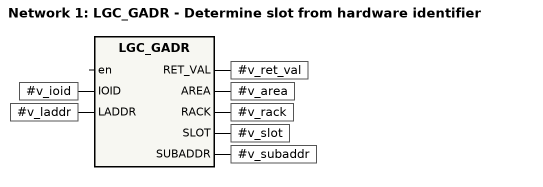
   #v_ret_val := LGC_GADR(IOID := #v_ioid,
                          LADDR := #v_laddr,
                          AREA => #v_area,
                          RACK => #v_rack,
                          SLOT => #v_slot,
                          SUBADDR => #v_subaddr);
END_REGION
END_FUNCTION_BLOCK

FUNCTION_BLOCK "FB_Fbd_ou001"   // FB169, FBD
{ S7_Optimized_Access := 'TRUE' }
   VAR_INPUT
      v_req : Bool;
      v_cont : Bool;
      v_len : UInt;
   END_VAR
   VAR_OUTPUT
      v_done : Bool;
      v_busy : Bool;
      v_error : Bool;
      v_status : Word;
   END_VAR
   VAR_IN_OUT
      v_connect : TCON_Param;
      v_data : Array[0..99] of Byte;
      v_com_rst : Bool;
      v_addr : Variant;
   END_VAR
   VAR
      inst : TSEND_C;
   END_VAR
BEGIN

REGION Network 1: TSEND_C - Send data via Ethernet
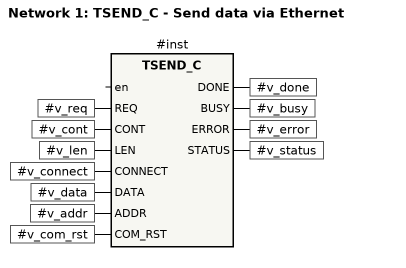
   #inst(REQ := #v_req,   // TSEND_C
         CONT := #v_cont,
         LEN := #v_len,
         CONNECT := #v_connect,
         DATA := #v_data,
         ADDR := #v_addr,
         COM_RST := #v_com_rst,
         DONE => #v_done,
         BUSY => #v_busy,
         ERROR => #v_error,
         STATUS => #v_status);
END_REGION
END_FUNCTION_BLOCK

FUNCTION_BLOCK "FB_Fbd_ou002"   // FB170, FBD
{ S7_Optimized_Access := 'TRUE' }
   VAR_INPUT
      v_req : Bool;
      v_cont : Bool;
      v_len : UDInt;
   END_VAR
   VAR_OUTPUT
      v_done : Bool;
      v_busy : Bool;
      v_error : Bool;
      v_status : Word;
   END_VAR
   VAR_IN_OUT
      v_connect : Array[0..99] of Byte;
      v_data : Array[0..99] of Byte;
      v_addr : Array[0..99] of Byte;
      v_com_rst : Bool;
   END_VAR
   VAR
      inst : TSEND_C;
   END_VAR
BEGIN

REGION Network 1: TSEND_C - Establishing a connection and sending data
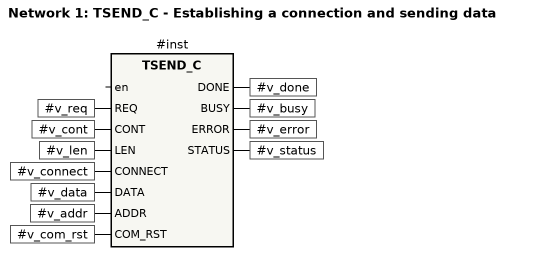
   #inst(REQ := #v_req,   // TSEND_C
         CONT := #v_cont,
         LEN := #v_len,
         CONNECT := #v_connect,
         DATA := #v_data,
         ADDR := #v_addr,
         COM_RST := #v_com_rst,
         DONE => #v_done,
         BUSY => #v_busy,
         ERROR => #v_error,
         STATUS => #v_status);
END_REGION
END_FUNCTION_BLOCK

FUNCTION_BLOCK "FB_Fbd_ou004"   // FB171, FBD
{ S7_Optimized_Access := 'TRUE' }
   VAR_INPUT
      v_en_r : Bool;
      v_cont : Bool;
      v_len : UDInt;
      v_adhoc : Bool;
   END_VAR
   VAR_OUTPUT
      v_done : Bool;
      v_busy : Bool;
      v_error : Bool;
      v_status : Word;
      v_rcvd_len : UDInt;
   END_VAR
   VAR_IN_OUT
      v_connect : Array[0..99] of Byte;
      v_data : Array[0..99] of Byte;
      v_addr : Array[0..99] of Byte;
      v_com_rst : Bool;
   END_VAR
   VAR
      inst : TRCV_C;
   END_VAR
BEGIN

REGION Network 1: TRCV_C - Establishing a connection and receiving data
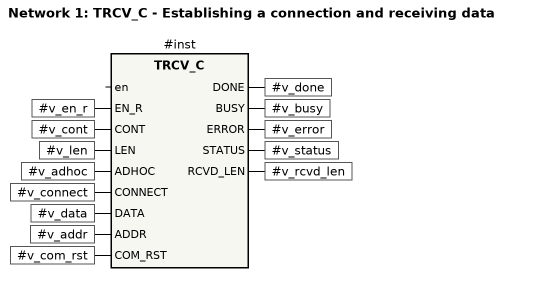
   #inst(EN_R := #v_en_r,   // TRCV_C
         CONT := #v_cont,
         LEN := #v_len,
         ADHOC := #v_adhoc,
         CONNECT := #v_connect,
         DATA := #v_data,
         ADDR := #v_addr,
         COM_RST := #v_com_rst,
         DONE => #v_done,
         BUSY => #v_busy,
         ERROR => #v_error,
         STATUS => #v_status,
         RCVD_LEN => #v_rcvd_len);
END_REGION
END_FUNCTION_BLOCK

FUNCTION_BLOCK "FB_Fbd_ou010"   // FB172, FBD
{ S7_Optimized_Access := 'TRUE' }
   VAR_INPUT
      v_req : Bool;
      v_id : Conn_Ouc;
   END_VAR
   VAR_OUTPUT
      v_done : Bool;
      v_busy : Bool;
      v_error : Bool;
      v_status : Word;
   END_VAR
   VAR_IN_OUT
      v_connect : TCON_Param;
   END_VAR
   VAR
      inst : TCON;
   END_VAR
BEGIN

REGION Network 1: TCON - Establish communication connection
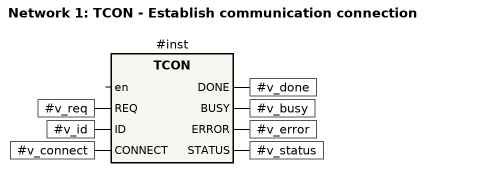
   #inst(REQ := #v_req,   // TCON
         ID := #v_id,
         CONNECT := #v_connect,
         DONE => #v_done,
         BUSY => #v_busy,
         ERROR => #v_error,
         STATUS => #v_status);
END_REGION
END_FUNCTION_BLOCK

FUNCTION_BLOCK "FB_Fbd_ou011"   // FB173, FBD
{ S7_Optimized_Access := 'TRUE' }
   VAR_INPUT
      v_req : Bool;
      v_id : Conn_Ouc;
   END_VAR
   VAR_OUTPUT
      v_done : Bool;
      v_busy : Bool;
      v_error : Bool;
      v_status : Word;
   END_VAR
   VAR_IN_OUT
      v_connect : Array[0..99] of Byte;
   END_VAR
   VAR
      inst : TCON;
   END_VAR
BEGIN

REGION Network 1: TCON - Establish communication connection
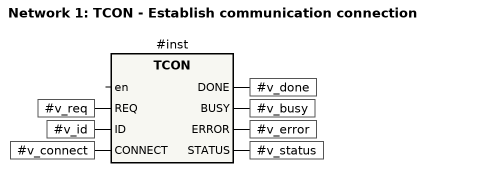
   #inst(REQ := #v_req,   // TCON
         ID := #v_id,
         CONNECT := #v_connect,
         DONE => #v_done,
         BUSY => #v_busy,
         ERROR => #v_error,
         STATUS => #v_status);
END_REGION
END_FUNCTION_BLOCK

FUNCTION_BLOCK "FB_Fbd_ou012"   // FB174, FBD
{ S7_Optimized_Access := 'TRUE' }
   VAR_INPUT
      v_req : Bool;
      v_id : Word;
   END_VAR
   VAR_OUTPUT
      v_done : Bool;
      v_busy : Bool;
      v_error : Bool;
      v_status : Word;
   END_VAR
   VAR
      inst : TDISCON;
   END_VAR
BEGIN

REGION Network 1: TDISCON - Terminate communication connection
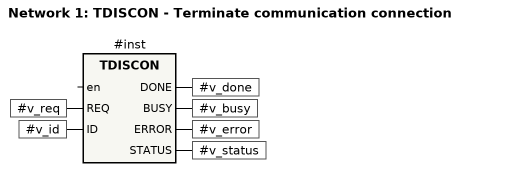
   #inst(REQ := #v_req, ID := #v_id, DONE => #v_done, BUSY => #v_busy, ERROR => #v_error, STATUS => #v_status);   // TDISCON
END_REGION
END_FUNCTION_BLOCK

FUNCTION_BLOCK "FB_Fbd_ou013"   // FB175, FBD
{ S7_Optimized_Access := 'TRUE' }
   VAR_INPUT
      v_req : Bool;
      v_id : Conn_Ouc;
      v_len : UInt;
   END_VAR
   VAR_OUTPUT
      v_done : Bool;
      v_busy : Bool;
      v_error : Bool;
      v_status : Word;
   END_VAR
   VAR_IN_OUT
      v_data : Array[0..99] of Byte;
   END_VAR
   VAR
      inst : TSEND;
   END_VAR
BEGIN

REGION Network 1: TSEND - Send data via communication connection
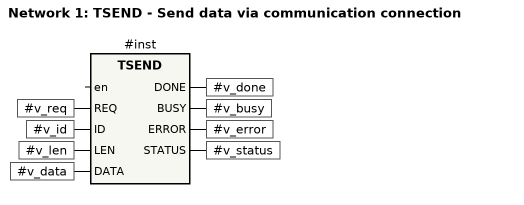
   #inst(REQ := #v_req,   // TSEND
         ID := #v_id,
         LEN := #v_len,
         DATA := #v_data,
         DONE => #v_done,
         BUSY => #v_busy,
         ERROR => #v_error,
         STATUS => #v_status);
END_REGION
END_FUNCTION_BLOCK

FUNCTION_BLOCK "FB_Fbd_ou014"   // FB176, FBD
{ S7_Optimized_Access := 'TRUE' }
   VAR_INPUT
      v_req : Bool;
      v_id : Conn_Ouc;
      v_len : UDInt;
   END_VAR
   VAR_OUTPUT
      v_done : Bool;
      v_busy : Bool;
      v_error : Bool;
      v_status : Word;
   END_VAR
   VAR_IN_OUT
      v_data : Array[0..99] of Byte;
   END_VAR
   VAR
      inst : TSEND;
   END_VAR
BEGIN

REGION Network 1: TSEND - Send data via communication connection
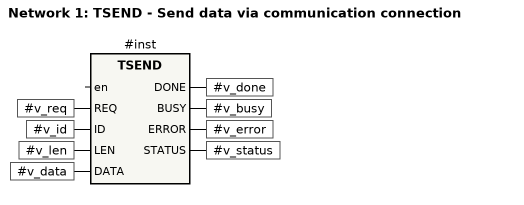
   #inst(REQ := #v_req,   // TSEND
         ID := #v_id,
         LEN := #v_len,
         DATA := #v_data,
         DONE => #v_done,
         BUSY => #v_busy,
         ERROR => #v_error,
         STATUS => #v_status);
END_REGION
END_FUNCTION_BLOCK

FUNCTION_BLOCK "FB_Fbd_ou016"   // FB177, FBD
{ S7_Optimized_Access := 'TRUE' }
   VAR_INPUT
      v_en_r : Bool;
      v_id : Conn_Ouc;
      v_len : UDInt;
      v_adhoc : Bool;
   END_VAR
   VAR_OUTPUT
      v_ndr : Bool;
      v_busy : Bool;
      v_error : Bool;
      v_status : Word;
      v_rcvd_len : UDInt;
   END_VAR
   VAR_IN_OUT
      v_data : Array[0..99] of Byte;
   END_VAR
   VAR
      inst : TRCV;
   END_VAR
BEGIN

REGION Network 1: TRCV - Receive data via communication connection
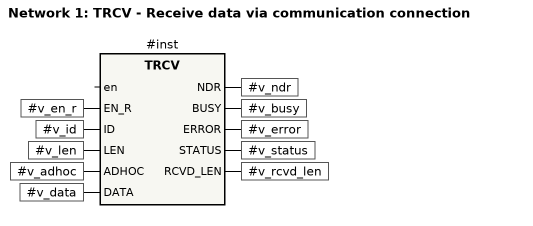
   #inst(EN_R := #v_en_r,   // TRCV
         ID := #v_id,
         LEN := #v_len,
         ADHOC := #v_adhoc,
         DATA := #v_data,
         NDR => #v_ndr,
         BUSY => #v_busy,
         ERROR => #v_error,
         STATUS => #v_status,
         RCVD_LEN => #v_rcvd_len);
END_REGION
END_FUNCTION_BLOCK

FUNCTION_BLOCK "FB_Fbd_ou017"   // FB178, FBD
{ S7_Optimized_Access := 'TRUE' }
   VAR_INPUT
      v_req : Bool;
      v_id : Conn_Ouc;
      v_len : UDInt;
   END_VAR
   VAR_OUTPUT
      v_done : Bool;
      v_busy : Bool;
      v_error : Bool;
      v_status : Word;
   END_VAR
   VAR_IN_OUT
      v_data : Array[0..99] of Byte;
      v_addr : Array[0..99] of Byte;
   END_VAR
   VAR
      inst : TUSEND;
   END_VAR
BEGIN

REGION Network 1: TUSEND - Sending data
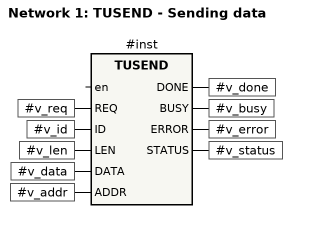
   #inst(REQ := #v_req,   // TUSEND
         ID := #v_id,
         LEN := #v_len,
         DATA := #v_data,
         ADDR := #v_addr,
         DONE => #v_done,
         BUSY => #v_busy,
         ERROR => #v_error,
         STATUS => #v_status);
END_REGION
END_FUNCTION_BLOCK

FUNCTION_BLOCK "FB_Fbd_ou018"   // FB179, FBD
{ S7_Optimized_Access := 'TRUE' }
   VAR_INPUT
      v_en_r : Bool;
      v_id : Conn_Ouc;
      v_len : UDInt;
   END_VAR
   VAR_OUTPUT
      v_ndr : Bool;
      v_error : Bool;
      v_busy : Bool;
      v_status : Word;
      v_rcvd_len : UDInt;
   END_VAR
   VAR_IN_OUT
      v_data : Array[0..99] of Byte;
      v_addr : Array[0..99] of Byte;
   END_VAR
   VAR
      inst : TURCV;
   END_VAR
BEGIN

REGION Network 1: TURCV - Receiving data
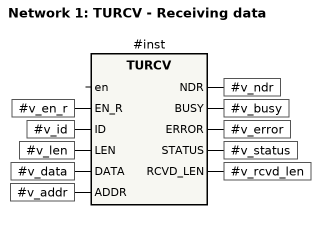
   #inst(EN_R := #v_en_r,   // TURCV
         ID := #v_id,
         LEN := #v_len,
         DATA := #v_data,
         ADDR := #v_addr,
         NDR => #v_ndr,
         BUSY => #v_busy,
         ERROR => #v_error,
         STATUS => #v_status,
         RCVD_LEN => #v_rcvd_len);
END_REGION
END_FUNCTION_BLOCK

FUNCTION_BLOCK "FB_Fbd_ou019"   // FB180, FBD
{ S7_Optimized_Access := 'TRUE' }
   VAR_INPUT
      v_req : Bool;
      v_id : Conn_Ouc;
   END_VAR
   VAR_OUTPUT
      v_done : Bool;
      v_busy : Bool;
      v_error : Bool;
      v_status : Word;
   END_VAR
   VAR
      inst : T_RESET;
   END_VAR
BEGIN

REGION Network 1: T_RESET - Resetting the connection
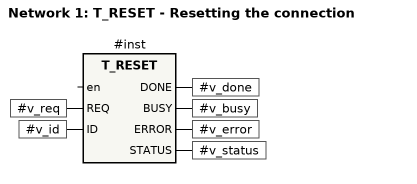
   #inst(REQ := #v_req, ID := #v_id, DONE => #v_done, BUSY => #v_busy, ERROR => #v_error, STATUS => #v_status);   // T_RESET
END_REGION
END_FUNCTION_BLOCK

FUNCTION_BLOCK "FB_Fbd_ou020"   // FB181, FBD
{ S7_Optimized_Access := 'TRUE' }
   VAR_INPUT
      v_req : Bool;
      v_id : Word;
   END_VAR
   VAR_OUTPUT
      v_done : Bool;
      v_busy : Bool;
      v_error : Bool;
      v_status : Word;
   END_VAR
   VAR_IN_OUT
      v_result : Array[0..99] of Byte;
   END_VAR
   VAR
      inst : T_DIAG;
   END_VAR
BEGIN

REGION Network 1: T_DIAG - Checking the connection
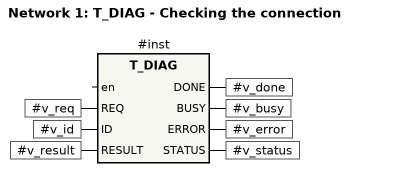
   #inst(REQ := #v_req,   // T_DIAG
         ID := #v_id,
         RESULT := #v_result,
         DONE => #v_done,
         BUSY => #v_busy,
         ERROR => #v_error,
         STATUS => #v_status);
END_REGION
END_FUNCTION_BLOCK

FUNCTION_BLOCK "FB_Fbd_sc003"   // FB182, FBD
{ S7_Optimized_Access := 'TRUE' }
   VAR_INPUT
      v_req : Bool;
      v_id : Conn_Prg;
      v_r_id : Conn_R_Id;
   END_VAR
   VAR_OUTPUT
      v_done : Bool;
      v_error : Bool;
      v_status : Word;
   END_VAR
   VAR_IN_OUT
      v_sd_1 : Variant;
      v_sd_2 : Variant;
      v_sd_3 : Variant;
      v_sd_4 : Variant;
   END_VAR
   VAR
      inst : USEND;
   END_VAR
BEGIN

REGION Network 1: USEND - Send data uncoordinated
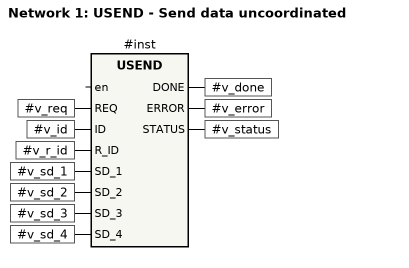
   #inst(REQ := #v_req,   // USEND
         ID := #v_id,
         R_ID := #v_r_id,
         SD_1 := #v_sd_1,
         SD_2 := #v_sd_2,
         SD_3 := #v_sd_3,
         SD_4 := #v_sd_4,
         DONE => #v_done,
         ERROR => #v_error,
         STATUS => #v_status);
END_REGION
END_FUNCTION_BLOCK

FUNCTION_BLOCK "FB_Fbd_sc004"   // FB183, FBD
{ S7_Optimized_Access := 'TRUE' }
   VAR_INPUT
      v_en_r : Bool;
      v_id : Conn_Prg;
      v_r_id : Conn_R_Id;
   END_VAR
   VAR_OUTPUT
      v_ndr : Bool;
      v_error : Bool;
      v_status : Word;
   END_VAR
   VAR_IN_OUT
      v_rd_1 : Variant;
      v_rd_2 : Variant;
      v_rd_3 : Variant;
      v_rd_4 : Variant;
   END_VAR
   VAR
      inst : URCV;
   END_VAR
BEGIN

REGION Network 1: URCV - Receive data uncoordinated
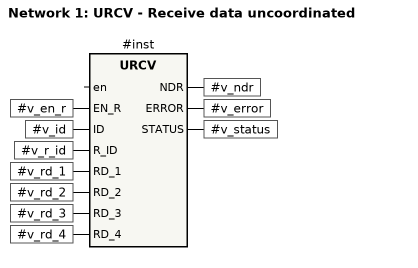
   #inst(EN_R := #v_en_r,   // URCV
         ID := #v_id,
         R_ID := #v_r_id,
         RD_1 := #v_rd_1,
         RD_2 := #v_rd_2,
         RD_3 := #v_rd_3,
         RD_4 := #v_rd_4,
         NDR => #v_ndr,
         ERROR => #v_error,
         STATUS => #v_status);
END_REGION
END_FUNCTION_BLOCK

FUNCTION_BLOCK "FB_Fbd_sc005"   // FB184, FBD
{ S7_Optimized_Access := 'TRUE' }
   VAR_INPUT
      v_req : Bool;
      v_r : Bool;
      v_id : Conn_Prg;
      v_r_id : Conn_R_Id;
   END_VAR
   VAR_OUTPUT
      v_done : Bool;
      v_error : Bool;
      v_status : Word;
   END_VAR
   VAR_IN_OUT
      v_sd_1 : Array[0..99] of Byte;
      v_len : Word;
   END_VAR
   VAR
      inst : BSEND;
   END_VAR
BEGIN

REGION Network 1: BSEND - Send data in segments
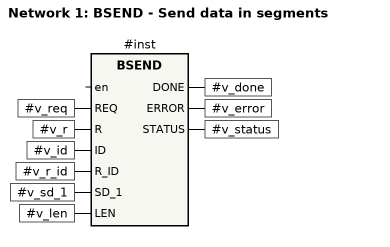
   #inst(REQ := #v_req,   // BSEND
         R := #v_r,
         ID := #v_id,
         R_ID := #v_r_id,
         SD_1 := #v_sd_1,
         LEN := #v_len,
         DONE => #v_done,
         ERROR => #v_error,
         STATUS => #v_status);
END_REGION
END_FUNCTION_BLOCK

FUNCTION_BLOCK "FB_Fbd_sc006"   // FB185, FBD
{ S7_Optimized_Access := 'TRUE' }
   VAR_INPUT
      v_en_r : Bool;
      v_id : Conn_Prg;
      v_r_id : Conn_R_Id;
   END_VAR
   VAR_OUTPUT
      v_ndr : Bool;
      v_error : Bool;
      v_status : Word;
   END_VAR
   VAR_IN_OUT
      v_rd_1 : Array[0..99] of Byte;
      v_len : Word;
   END_VAR
   VAR
      inst : BRCV;
   END_VAR
BEGIN

REGION Network 1: BRCV - Receive data in segments
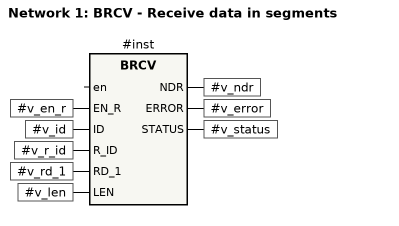
   #inst(EN_R := #v_en_r,   // BRCV
         ID := #v_id,
         R_ID := #v_r_id,
         RD_1 := #v_rd_1,
         LEN := #v_len,
         NDR => #v_ndr,
         ERROR => #v_error,
         STATUS => #v_status);
END_REGION
END_FUNCTION_BLOCK

FUNCTION_BLOCK "FB_Scl_sl041"   // FB186, SCL
{ S7_Optimized_Access := 'TRUE' }
VERSION : 0.1
   VAR_INPUT
      v_in : Array[0..9] of Date;
      v_count : USInt;
   END_VAR
   VAR_OUTPUT
      v_out : Array[0..9] of Date;
   END_VAR
BEGIN
   MOVE_BLK(IN := #v_in[0], COUNT := #v_count, OUT => #v_out[0]);
END_FUNCTION_BLOCK

FUNCTION_BLOCK "FB_Scl_sl047"   // FB187, SCL
{ S7_Optimized_Access := 'TRUE' }
VERSION : 0.1
   VAR_INPUT
      v_in : Array[0..9] of Byte;
      v_count_in : USInt;
   END_VAR
   VAR_OUTPUT
      v_out : Array[0..9] of Bool;
   END_VAR
BEGIN
   SCATTER_BLK(IN := #v_in[0], COUNT_IN := #v_count_in, OUT => #v_out[0]);
END_FUNCTION_BLOCK

FUNCTION_BLOCK "FB_Scl_sl043"   // FB188, SCL
{ S7_Optimized_Access := 'TRUE' }
VERSION : 0.1
   VAR_INPUT
      v_in : Array[0..9] of Date;
      v_count : USInt;
   END_VAR
   VAR_OUTPUT
      v_out : Array[0..9] of Date;
   END_VAR
BEGIN
   UMOVE_BLK(IN := #v_in[0], COUNT := #v_count, OUT => #v_out[0]);
END_FUNCTION_BLOCK

FUNCTION_BLOCK "FB_Scl_sl049"   // FB189, SCL
{ S7_Optimized_Access := 'TRUE' }
VERSION : 0.1
   VAR_INPUT
      v_in : Array[0..9] of Bool;
      v_count_out : USInt;
   END_VAR
   VAR_OUTPUT
      v_out : Array[0..9] of Byte;
   END_VAR
BEGIN
   GATHER_BLK(IN := #v_in[0], COUNT_OUT := #v_count_out, OUT => #v_out[0]);
END_FUNCTION_BLOCK

FUNCTION_BLOCK "FB_Scl_sl103"   // FB190, SCL
{ S7_Optimized_Access := 'TRUE' }
VERSION : 0.1
   VAR_INPUT
      v_in : UInt;
   END_VAR
   VAR_OUTPUT
      v_ret : UInt;
   END_VAR
BEGIN
   #v_ret := DECO(IN := #v_in);
END_FUNCTION_BLOCK

FUNCTION_BLOCK "FB_Scl_sl104"   // FB191, SCL
{ S7_Optimized_Access := 'TRUE' }
VERSION : 0.1
   VAR_INPUT
      v_in : Word;
   END_VAR
   VAR_OUTPUT
      v_ret : Word;
   END_VAR
BEGIN
   #v_ret := ENCO(IN := #v_in);
END_FUNCTION_BLOCK

FUNCTION_BLOCK "FB_Scl_sl108"   // FB192, SCL
{ S7_Optimized_Access := 'TRUE' }
VERSION : 0.1
   VAR_INPUT
      v_in : Word;
      v_n : USInt;
   END_VAR
   VAR_OUTPUT
      v_ret : Word;
   END_VAR
BEGIN
   #v_ret := SHR(IN := #v_in, N := #v_n);
END_FUNCTION_BLOCK

FUNCTION_BLOCK "FB_Scl_sl109"   // FB193, SCL
{ S7_Optimized_Access := 'TRUE' }
VERSION : 0.1
   VAR_INPUT
      v_in : Word;
      v_n : USInt;
   END_VAR
   VAR_OUTPUT
      v_ret : Word;
   END_VAR
BEGIN
   #v_ret := SHL(IN := #v_in, N := #v_n);
END_FUNCTION_BLOCK

FUNCTION_BLOCK "FB_Scl_sl110"   // FB194, SCL
{ S7_Optimized_Access := 'TRUE' }
VERSION : 0.1
   VAR_INPUT
      v_in : Word;
      v_n : USInt;
   END_VAR
   VAR_OUTPUT
      v_ret : Word;
   END_VAR
BEGIN
   #v_ret := ROR(IN := #v_in, N := #v_n);
END_FUNCTION_BLOCK

FUNCTION_BLOCK "FB_Scl_sl111"   // FB195, SCL
{ S7_Optimized_Access := 'TRUE' }
VERSION : 0.1
   VAR_INPUT
      v_in : Word;
      v_n : USInt;
   END_VAR
   VAR_OUTPUT
      v_ret : Word;
   END_VAR
BEGIN
   #v_ret := ROL(IN := #v_in, N := #v_n);
END_FUNCTION_BLOCK

FUNCTION_BLOCK "FB_Scl_sl112"   // FB196, SCL
{ S7_Optimized_Access := 'TRUE' }
VERSION : 0.1
   VAR_INPUT
      v_reset : Bool;
      v_jog : Bool;
      v_drum_en : Bool;
      v_lst_step : Byte;
   END_VAR
   VAR_OUTPUT
      v_q : Bool;
      v_out_word : Word;
      v_err_code : Word;
   END_VAR
   VAR
      inst : DRUM;
   END_VAR
BEGIN
   #inst(RESET := #v_reset, JOG := #v_jog, DRUM_EN := #v_drum_en, LST_STEP := #v_lst_step, Q => #v_q, OUT_WORD => #v_out_word, ERR_CODE => #v_err_code);
END_FUNCTION_BLOCK

FUNCTION_BLOCK "FB_Scl_sl113"   // FB197, SCL
{ S7_Optimized_Access := 'TRUE' }
VERSION : 0.1
   VAR_INPUT
      v_cmd : Bool;
      v_o_fb : Bool;
      v_c_fb : Bool;
   END_VAR
   VAR_OUTPUT
      v_q : Bool;
      v_oa : Bool;
      v_ca : Bool;
   END_VAR
   VAR
      inst : DCAT;
   END_VAR
BEGIN
   #inst(CMD := #v_cmd, O_FB := #v_o_fb, C_FB := #v_c_fb, Q => #v_q, OA => #v_oa, CA => #v_ca);
END_FUNCTION_BLOCK

FUNCTION_BLOCK "FB_Scl_sl114"   // FB198, SCL
{ S7_Optimized_Access := 'TRUE' }
VERSION : 0.1
   VAR_INPUT
      v_o_cmd : Bool;
      v_c_cmd : Bool;
      v_s_cmd : Bool;
      v_o_fb : Bool;
      v_c_fb : Bool;
   END_VAR
   VAR_OUTPUT
      v_oo : Bool;
      v_co : Bool;
      v_oa : Bool;
      v_ca : Bool;
      v_q : Bool;
   END_VAR
   VAR
      inst : MCAT;
   END_VAR
BEGIN
   #inst(O_CMD := #v_o_cmd, C_CMD := #v_c_cmd, S_CMD := #v_s_cmd, O_FB := #v_o_fb, C_FB := #v_c_fb, OO => #v_oo, CO => #v_co, OA => #v_oa, CA => #v_ca, Q => #v_q);
END_FUNCTION_BLOCK

FUNCTION_BLOCK "FB_Scl_sl115"   // FB199, SCL
{ S7_Optimized_Access := 'TRUE' }
VERSION : 0.1
   VAR_INPUT
      v_in_bit0 : Bool;
      v_in_bit1 : Bool;
      v_in_bit2 : Bool;
      v_in_bit3 : Bool;
      v_in_bit4 : Bool;
      v_in_bit5 : Bool;
      v_in_bit6 : Bool;
      v_in_bit7 : Bool;
      v_in_bit8 : Bool;
      v_in_bit9 : Bool;
      v_in_bit10 : Bool;
      v_in_bit11 : Bool;
      v_in_bit12 : Bool;
      v_in_bit13 : Bool;
      v_in_bit14 : Bool;
      v_in_bit15 : Bool;
      v_cmp_step : Byte;
   END_VAR
   VAR_OUTPUT
      v_out : Bool;
      v_err_code : Word;
   END_VAR
   VAR
      inst : IMC;
   END_VAR
BEGIN
   #inst(IN_BIT0 := #v_in_bit0, IN_BIT1 := #v_in_bit1, IN_BIT2 := #v_in_bit2, IN_BIT3 := #v_in_bit3, IN_BIT4 := #v_in_bit4, IN_BIT5 := #v_in_bit5, IN_BIT6 := #v_in_bit6, IN_BIT7 := #v_in_bit7, IN_BIT8 := #v_in_bit8, IN_BIT9 := #v_in_bit9, IN_BIT10 := #v_in_bit10, IN_BIT11 := #v_in_bit11, IN_BIT12 := #v_in_bit12, IN_BIT13 := #v_in_bit13, IN_BIT14 := #v_in_bit14, IN_BIT15 := #v_in_bit15, CMP_STEP := #v_cmp_step, OUT => #v_out, ERR_CODE => #v_err_code);
END_FUNCTION_BLOCK

FUNCTION_BLOCK "FB_Scl_sl116"   // FB203, SCL
{ S7_Optimized_Access := 'TRUE' }
VERSION : 0.1
   VAR_INPUT
      v_in_bit0 : Bool;
      v_in_bit1 : Bool;
      v_in_bit2 : Bool;
      v_in_bit3 : Bool;
      v_in_bit4 : Bool;
      v_in_bit5 : Bool;
      v_in_bit6 : Bool;
      v_in_bit7 : Bool;
      v_in_bit8 : Bool;
      v_in_bit9 : Bool;
      v_in_bit10 : Bool;
      v_in_bit11 : Bool;
      v_in_bit12 : Bool;
      v_in_bit13 : Bool;
      v_in_bit14 : Bool;
      v_in_bit15 : Bool;
   END_VAR
   VAR_OUTPUT
      v_out : Bool;
      v_out_step : Byte;
      v_err_code : Word;
   END_VAR
   VAR
      inst : SMC;
   END_VAR
BEGIN
   #inst(IN_BIT0 := #v_in_bit0, IN_BIT1 := #v_in_bit1, IN_BIT2 := #v_in_bit2, IN_BIT3 := #v_in_bit3, IN_BIT4 := #v_in_bit4, IN_BIT5 := #v_in_bit5, IN_BIT6 := #v_in_bit6, IN_BIT7 := #v_in_bit7, IN_BIT8 := #v_in_bit8, IN_BIT9 := #v_in_bit9, IN_BIT10 := #v_in_bit10, IN_BIT11 := #v_in_bit11, IN_BIT12 := #v_in_bit12, IN_BIT13 := #v_in_bit13, IN_BIT14 := #v_in_bit14, IN_BIT15 := #v_in_bit15, OUT => #v_out, OUT_STEP => #v_out_step, ERR_CODE => #v_err_code);
END_FUNCTION_BLOCK

FUNCTION_BLOCK "FB_Scl_sl117"   // FB205, SCL
{ S7_Optimized_Access := 'TRUE' }
VERSION : 0.1
   VAR_INPUT
      v_in : Real;
      v_sample_t : Int;
   END_VAR
   VAR_OUTPUT
      v_out : Real;
      v_err_code : Word;
   END_VAR
   VAR
      inst : LEAD_LAG;
   END_VAR
BEGIN
   #inst(IN := #v_in, SAMPLE_T := #v_sample_t, OUT => #v_out, ERR_CODE => #v_err_code);
END_FUNCTION_BLOCK

FUNCTION_BLOCK "FB_Scl_sl118"   // FB207, SCL
{ S7_Optimized_Access := 'TRUE' }
VERSION : 0.1
   VAR_INPUT
      v_in : Word;
   END_VAR
   VAR_OUTPUT
      v_out : DWord;
   END_VAR
BEGIN
   SEG(IN := #v_in, OUT => #v_out);
END_FUNCTION_BLOCK

FUNCTION_BLOCK "FB_Scl_sl119"   // FB208, SCL
{ S7_Optimized_Access := 'TRUE' }
VERSION : 0.1
   VAR_INPUT
      v_in : Word;
   END_VAR
   VAR_OUTPUT
      v_ret : Word;
   END_VAR
BEGIN
   #v_ret := BCDCPL(IN := #v_in);
END_FUNCTION_BLOCK

FUNCTION_BLOCK "FB_Scl_sl120"   // FB209, SCL
{ S7_Optimized_Access := 'TRUE' }
VERSION : 0.1
   VAR_INPUT
      v_in : DWord;
   END_VAR
   VAR_OUTPUT
      v_ret : DWord;
   END_VAR
BEGIN
   #v_ret := BITSUM(IN := #v_in);
END_FUNCTION_BLOCK

FUNCTION_BLOCK "FB_Lad_ex159"   // FB210, LAD
{ S7_Optimized_Access := 'TRUE' }
   VAR_INPUT
      v_ioid : Byte;
      v_laddr : Hw_Any;
   END_VAR
   VAR_OUTPUT
      v_ret_val : Int;
      v_pecount : Int;
      v_pacount : Int;
   END_VAR
BEGIN

REGION Network 1: RD_LGADR - Determine IO addresses from the hardware identifier
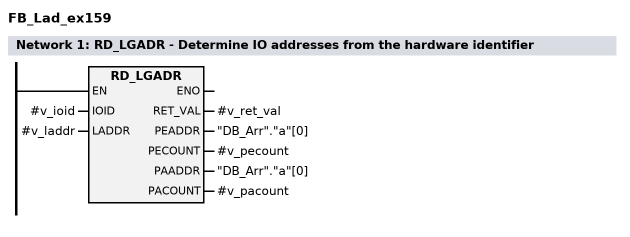
   #v_ret_val := RD_LGADR(IOID := #v_ioid,
                          LADDR := #v_laddr,
                          PEADDR => "DB_Arr"."a"[0],
                          PECOUNT => #v_pecount,
                          PAADDR => "DB_Arr"."a"[0],
                          PACOUNT => #v_pacount);
END_REGION
END_FUNCTION_BLOCK

FUNCTION_BLOCK "FX_Fbd_ex003"   // FB211, FBD
{ S7_Optimized_Access := 'TRUE' }
VERSION : 0.1
   VAR_INPUT
      "a" : Bool;
      "b" : Bool;
      c : Bool;
      ia : Int;
      ib : Int;
      ic : Int;
      da : DInt;
      db : DInt;
      ra : Real;
      rb : Real;
      wa : Word;
      wb : Word;
      dwa : DWord;
      ba : Byte;
      ta : Time;
      tb : Time;
      s1 : String;
      s2 : String;
   END_VAR
   VAR_OUTPUT
      q : Bool;
      q2 : Bool;
      io : Int;
      io2 : Int;
      dout : DInt;
      rout : Real;
      wout : Word;
      dwout : DWord;
      bout : Byte;
      tout : Time;
      sout : String;
   END_VAR
   VAR_IN_OUT
      x_time : Time;
      arr : Array[0..9] of Int;
      barr : Array[0..7] of Bool;
      iinout : Int;
   END_VAR
   VAR
      ton1 : TON_TIME;
      tof1 : TOF_TIME;
      tp1 : TP_TIME;
      tonr1 : TONR_TIME;
      ctu1 : CTU_INT;
      ctd1 : CTD_INT;
      ctud1 : CTUD_INT;
      rtrig1 : R_TRIG;
      ftrig1 : F_TRIG;
      edge1 : Bool;
      edge2 : Bool;
      stat1 : Bool;
      stat2 : Bool;
      stati : Int;
   END_VAR
   VAR_TEMP
      t1 : Bool;
      t2 : Bool;
      ti : Int;
      td : DInt;
      tr : Real;
      tw : Word;
      tt : Time;
      var1 : Variant;
   END_VAR
BEGIN

REGION Network 1: ---| |--- - Normally open contact
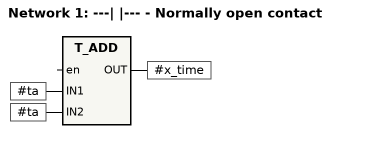
   #x_time := T_ADD(IN1 := #ta, IN2 := #ta);
END_REGION
END_FUNCTION_BLOCK

FUNCTION_BLOCK "FX_Fbd_ex004"   // FB212, FBD
{ S7_Optimized_Access := 'TRUE' }
VERSION : 0.1
   VAR_INPUT
      "a" : Bool;
      "b" : Bool;
      c : Bool;
      ia : Int;
      ib : Int;
      ic : Int;
      da : DInt;
      db : DInt;
      ra : Real;
      rb : Real;
      wa : Word;
      wb : Word;
      dwa : DWord;
      ba : Byte;
      ta : Time;
      tb : Time;
      s1 : String;
      s2 : String;
   END_VAR
   VAR_OUTPUT
      q : Bool;
      q2 : Bool;
      io : Int;
      io2 : Int;
      dout : DInt;
      rout : Real;
      wout : Word;
      dwout : DWord;
      bout : Byte;
      tout : Time;
      sout : String;
   END_VAR
   VAR_IN_OUT
      x_time : Time;
      arr : Array[0..9] of Int;
      barr : Array[0..7] of Bool;
      iinout : Int;
   END_VAR
   VAR
      ton1 : TON_TIME;
      tof1 : TOF_TIME;
      tp1 : TP_TIME;
      tonr1 : TONR_TIME;
      ctu1 : CTU_INT;
      ctd1 : CTD_INT;
      ctud1 : CTUD_INT;
      rtrig1 : R_TRIG;
      ftrig1 : F_TRIG;
      edge1 : Bool;
      edge2 : Bool;
      stat1 : Bool;
      stat2 : Bool;
      stati : Int;
   END_VAR
   VAR_TEMP
      t1 : Bool;
      t2 : Bool;
      ti : Int;
      td : DInt;
      tr : Real;
      tw : Word;
      tt : Time;
      var1 : Variant;
   END_VAR
BEGIN

REGION Network 1: ---| |--- - Normally open contact
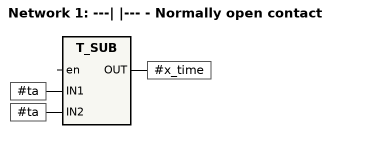
   #x_time := T_SUB(IN1 := #ta, IN2 := #ta);
END_REGION
END_FUNCTION_BLOCK

FUNCTION_BLOCK "FX_Fbd_ex018"   // FB213, FBD
{ S7_Optimized_Access := 'TRUE' }
VERSION : 0.1
   VAR_INPUT
      "a" : Bool;
      "b" : Bool;
      c : Bool;
      ia : Int;
      ib : Int;
      ic : Int;
      da : DInt;
      db : DInt;
      ra : Real;
      rb : Real;
      wa : Word;
      wb : Word;
      dwa : DWord;
      ba : Byte;
      ta : Time;
      tb : Time;
      s1 : String;
      s2 : String;
   END_VAR
   VAR_OUTPUT
      q : Bool;
      q2 : Bool;
      io : Int;
      io2 : Int;
      dout : DInt;
      rout : Real;
      wout : Word;
      dwout : DWord;
      bout : Byte;
      tout : Time;
      sout : String;
   END_VAR
   VAR_IN_OUT
      arr : Array[0..9] of Int;
      barr : Array[0..7] of Bool;
      iinout : Int;
   END_VAR
   VAR
      ton1 : TON_TIME;
      tof1 : TOF_TIME;
      tp1 : TP_TIME;
      tonr1 : TONR_TIME;
      ctu1 : CTU_INT;
      ctd1 : CTD_INT;
      ctud1 : CTUD_INT;
      rtrig1 : R_TRIG;
      ftrig1 : F_TRIG;
      edge1 : Bool;
      edge2 : Bool;
      stat1 : Bool;
      stat2 : Bool;
      stati : Int;
   END_VAR
   VAR_TEMP
      t1 : Bool;
      t2 : Bool;
      ti : Int;
      td : DInt;
      tr : Real;
      tw : Word;
      tt : Time;
      var1 : Variant;
   END_VAR
BEGIN

REGION Network 1: ---| |--- - Normally open contact
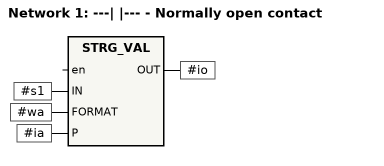
   STRG_VAL(IN := #s1, FORMAT := #wa, P := #ia, OUT => #io);
END_REGION
END_FUNCTION_BLOCK

FUNCTION_BLOCK "FX_Fbd_ex019"   // FB214, FBD
{ S7_Optimized_Access := 'TRUE' }
VERSION : 0.1
   VAR_INPUT
      "a" : Bool;
      "b" : Bool;
      c : Bool;
      ia : Int;
      ib : Int;
      ic : Int;
      da : DInt;
      db : DInt;
      ra : Real;
      rb : Real;
      wa : Word;
      wb : Word;
      dwa : DWord;
      ba : Byte;
      ta : Time;
      tb : Time;
      s1 : String;
      s2 : String;
   END_VAR
   VAR_OUTPUT
      q : Bool;
      q2 : Bool;
      io : Int;
      io2 : Int;
      dout : DInt;
      rout : Real;
      wout : Word;
      dwout : DWord;
      bout : Byte;
      tout : Time;
      sout : String;
   END_VAR
   VAR_IN_OUT
      arr : Array[0..9] of Int;
      barr : Array[0..7] of Bool;
      iinout : Int;
   END_VAR
   VAR
      ton1 : TON_TIME;
      tof1 : TOF_TIME;
      tp1 : TP_TIME;
      tonr1 : TONR_TIME;
      ctu1 : CTU_INT;
      ctd1 : CTD_INT;
      ctud1 : CTUD_INT;
      rtrig1 : R_TRIG;
      ftrig1 : F_TRIG;
      edge1 : Bool;
      edge2 : Bool;
      stat1 : Bool;
      stat2 : Bool;
      stati : Int;
   END_VAR
   VAR_TEMP
      t1 : Bool;
      t2 : Bool;
      ti : Int;
      td : DInt;
      tr : Real;
      tw : Word;
      tt : Time;
      var1 : Variant;
   END_VAR
BEGIN

REGION Network 1: ---| |--- - Normally open contact
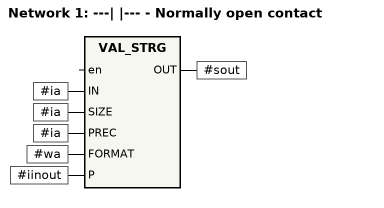
   VAL_STRG(IN := #ia, SIZE := #ia, PREC := #ia, FORMAT := #wa, P := #iinout, OUT => #sout);
END_REGION
END_FUNCTION_BLOCK

FUNCTION_BLOCK "FX_Fbd_ex021"   // FB215, FBD
{ S7_Optimized_Access := 'TRUE' }
VERSION : 0.1
   VAR_INPUT
      "a" : Bool;
      "b" : Bool;
      c : Bool;
      ia : Int;
      ib : Int;
      ic : Int;
      da : DInt;
      db : DInt;
      ra : Real;
      rb : Real;
      wa : Word;
      wb : Word;
      dwa : DWord;
      ba : Byte;
      ta : Time;
      tb : Time;
      s1 : String;
      s2 : String;
   END_VAR
   VAR_OUTPUT
      q : Bool;
      q2 : Bool;
      io : Int;
      io2 : Int;
      dout : DInt;
      rout : Real;
      wout : Word;
      dwout : DWord;
      bout : Byte;
      tout : Time;
      sout : String;
   END_VAR
   VAR_IN_OUT
      x_variant : Variant;
      arr : Array[0..9] of Int;
      barr : Array[0..7] of Bool;
      iinout : Int;
   END_VAR
   VAR
      ton1 : TON_TIME;
      tof1 : TOF_TIME;
      tp1 : TP_TIME;
      tonr1 : TONR_TIME;
      ctu1 : CTU_INT;
      ctd1 : CTD_INT;
      ctud1 : CTUD_INT;
      rtrig1 : R_TRIG;
      ftrig1 : F_TRIG;
      edge1 : Bool;
      edge2 : Bool;
      stat1 : Bool;
      stat2 : Bool;
      stati : Int;
   END_VAR
   VAR_TEMP
      t1 : Bool;
      t2 : Bool;
      ti : Int;
      td : DInt;
      tr : Real;
      tw : Word;
      tt : Time;
      var1 : Variant;
   END_VAR
BEGIN

REGION Network 1: ---| |--- - Normally open contact
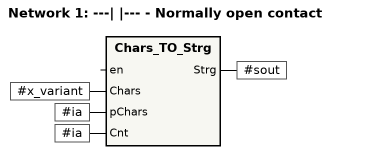
   // no SCL statement known for Chars_TO_Strg: written as a call
   Chars_TO_Strg(Chars := #x_variant, pChars := #ia, Cnt := #ia, Strg => #sout);
END_REGION
END_FUNCTION_BLOCK

FUNCTION_BLOCK "FX_Fbd_ex027"   // FB216, FBD
{ S7_Optimized_Access := 'TRUE' }
VERSION : 0.1
   VAR_INPUT
      "a" : Bool;
      "b" : Bool;
      c : Bool;
      ia : Int;
      ib : Int;
      ic : Int;
      da : DInt;
      db : DInt;
      ra : Real;
      rb : Real;
      wa : Word;
      wb : Word;
      dwa : DWord;
      ba : Byte;
      ta : Time;
      tb : Time;
      s1 : String;
      s2 : String;
   END_VAR
   VAR_OUTPUT
      q : Bool;
      q2 : Bool;
      io : Int;
      io2 : Int;
      dout : DInt;
      rout : Real;
      wout : Word;
      dwout : DWord;
      bout : Byte;
      tout : Time;
      sout : String;
   END_VAR
   VAR_IN_OUT
      arr : Array[0..9] of Int;
      barr : Array[0..7] of Bool;
      iinout : Int;
   END_VAR
   VAR
      ton1 : TON_TIME;
      tof1 : TOF_TIME;
      tp1 : TP_TIME;
      tonr1 : TONR_TIME;
      ctu1 : CTU_INT;
      ctd1 : CTD_INT;
      ctud1 : CTUD_INT;
      rtrig1 : R_TRIG;
      ftrig1 : F_TRIG;
      edge1 : Bool;
      edge2 : Bool;
      stat1 : Bool;
      stat2 : Bool;
      stati : Int;
   END_VAR
   VAR_TEMP
      t1 : Bool;
      t2 : Bool;
      ti : Int;
      td : DInt;
      tr : Real;
      tw : Word;
      tt : Time;
      var1 : Variant;
   END_VAR
BEGIN

REGION Network 1: ---| |--- - Normally open contact
